Yaskawa INFORM job: cattua0.JBI

/JOB
//NAME cattua0
//POS
///NPOS 130,0,0,0,0,0
///TOOL 9
///POSTYPE PULSE
///PULSE
C00000=-149478,-3800,-72601,-72634,-83747,-23013
C00001=-158362,27238,-42051,-68147,-87155,-20871
C00002=-155378,40422,-20095,-70093,-86314,-22222
C00003=-152934,54036,4519,-71957,-85739,-23985
C00004=-152872,54426,5251,-72009,-85726,-24041
C00005=-152818,54830,6002,-72058,-85717,-24097
C00006=-152775,55247,6768,-72103,-85712,-24152
C00007=-152741,55675,7548,-72144,-85712,-24206
C00008=-152718,56112,8337,-72182,-85717,-24260
C00009=-152706,56556,9133,-72216,-85727,-24313
C00010=-152703,57006,9933,-72246,-85742,-24364
C00011=-152712,57461,10733,-72271,-85762,-24415
C00012=-152730,57917,11532,-72293,-85786,-24464
C00013=-152759,58374,12326,-72310,-85815,-24511
C00014=-152798,58830,13113,-72324,-85848,-24557
C00015=-152846,59283,13889,-72334,-85886,-24600
C00016=-152903,59731,14652,-72340,-85927,-24642
C00017=-152969,60172,15400,-72342,-85973,-24683
C00018=-153124,61027,16837,-72336,-86074,-24757
C00019=-153307,61842,18195,-72317,-86186,-24823
C00020=-153524,62645,19517,-72286,-86315,-24883
C00021=-153773,63424,20787,-72241,-86458,-24938
C00022=-154052,64166,21985,-72184,-86615,-24985
C00023=-154358,64860,23092,-72114,-86783,-25024
C00024=-154687,65495,24091,-72033,-86960,-25055
C00025=-155034,66063,24971,-71941,-87145,-25077
C00026=-155395,66557,25719,-71839,-87334,-25089
C00027=-156090,67486,27164,-71650,-87700,-25120
C00028=-156792,68395,28628,-71464,-88074,-25159
C00029=-157502,69283,30109,-71285,-88455,-25207
C00030=-158217,70146,31604,-71111,-88843,-25263
C00031=-158938,70984,33108,-70945,-89238,-25327
C00032=-159661,71794,34620,-70786,-89640,-25400
C00033=-160387,72575,36134,-70636,-90046,-25480
C00034=-161114,73326,37650,-70495,-90458,-25569
C00035=-161841,74047,39164,-70364,-90874,-25665
C00036=-162568,74735,40675,-70242,-91293,-25769
C00037=-163292,75392,42179,-70132,-91716,-25881
C00038=-164013,76015,43673,-70033,-92142,-25999
C00039=-164729,76606,45157,-69946,-92569,-26124
C00040=-165440,77164,46627,-69871,-92997,-26256
C00041=-166143,77688,48082,-69808,-93425,-26393
C00042=-166839,78181,49519,-69758,-93852,-26537
C00043=-167197,78385,50174,-69730,-94071,-26606
C00044=-167566,78510,50675,-69688,-94290,-26661
C00045=-167940,78553,51011,-69632,-94507,-26702
C00046=-168316,78512,51178,-69562,-94720,-26728
C00047=-168690,78390,51174,-69478,-94926,-26737
C00048=-169057,78191,51002,-69380,-95123,-26731
C00049=-169413,77920,50673,-69271,-95307,-26709
C00050=-169759,77583,50193,-69149,-95480,-26672
C00051=-170104,77167,49544,-69010,-95646,-26618
C00052=-170444,76676,48726,-68854,-95801,-26547
C00053=-170773,76114,47744,-68684,-95944,-26458
C00054=-170932,75809,47195,-68593,-96010,-26408
C00055=-171087,75489,46610,-68500,-96071,-26354
C00056=-171237,75156,45990,-68403,-96128,-26295
C00057=-171381,74810,45337,-68304,-96181,-26234
C00058=-171519,74454,44656,-68203,-96228,-26168
C00059=-171651,74088,43948,-68101,-96271,-26100
C00060=-171776,73715,43217,-67997,-96308,-26029
C00061=-171893,73336,42467,-67892,-96340,-25956
C00062=-172106,72568,40924,-67682,-96388,-25804
C00063=-176209,59482,15170,-63884,-97305,-23273
C00064=-180964,47935,-6371,-60041,-98451,-21150
C00065=-181093,47637,-6920,-59937,-98479,-21095
C00066=-181207,47321,-7519,-59832,-98497,-21036
C00067=-181305,46992,-8163,-59728,-98503,-20972
C00068=-181384,46655,-8839,-59627,-98496,-20905
C00069=-181443,46314,-9539,-59531,-98477,-20837
C00070=-181482,45976,-10249,-59441,-98446,-20767
C00071=-181498,45645,-10960,-59360,-98405,-20698
C00072=-181495,45326,-11657,-59288,-98354,-20632
C00073=-181473,45023,-12333,-59226,-98295,-20567
C00074=-181431,44725,-13010,-59171,-98226,-20504
C00075=-181369,44435,-13683,-59126,-98148,-20441
C00076=-181287,44157,-14341,-59090,-98061,-20381
C00077=-181186,43895,-14975,-59065,-97966,-20324
C00078=-181067,43652,-15576,-59051,-97865,-20271
C00079=-180931,43432,-16137,-59049,-97758,-20223
C00080=-180781,43237,-16651,-59058,-97649,-20180
C00081=-180331,42715,-18030,-59105,-97335,-20069
C00082=-179870,42191,-19389,-59167,-97022,-19965
C00083=-179397,41663,-20725,-59243,-96709,-19868
C00084=-178913,41133,-22039,-59333,-96396,-19778
C00085=-178417,40599,-23328,-59437,-96085,-19694
C00086=-177910,40063,-24592,-59555,-95774,-19618
C00087=-177391,39523,-25830,-59686,-95465,-19550
C00088=-176861,38981,-27041,-59831,-95157,-19488
C00089=-176321,38437,-28225,-59989,-94850,-19434
C00090=-175769,37891,-29380,-60160,-94545,-19387
C00091=-175207,37342,-30505,-60344,-94242,-19347
C00092=-174635,36792,-31599,-60540,-93941,-19315
C00093=-174053,36240,-32663,-60748,-93641,-19290
C00094=-173462,35687,-33694,-60968,-93344,-19272
C00095=-172862,35132,-34693,-61198,-93049,-19262
C00096=-172252,34577,-35659,-61440,-92755,-19259
C00097=-171634,34021,-36591,-61692,-92464,-19263
C00098=-171008,33464,-37488,-61954,-92175,-19274
C00099=-170375,32907,-38351,-62225,-91888,-19293
C00100=-169734,32350,-39178,-62506,-91604,-19319
C00101=-169086,31793,-39970,-62795,-91321,-19352
C00102=-168432,31237,-40725,-63091,-91041,-19392
C00103=-167773,30682,-41443,-63396,-90762,-19440
C00104=-167108,30129,-42124,-63707,-90486,-19494
C00105=-166440,29577,-42767,-64025,-90212,-19555
C00106=-165767,29028,-43372,-64348,-89940,-19622
C00107=-165092,28481,-43940,-64676,-89670,-19697
C00108=-164414,27937,-44469,-65009,-89403,-19777
C00109=-163734,27396,-44960,-65345,-89137,-19864
C00110=-163053,26860,-45412,-65685,-88873,-19957
C00111=-162372,26328,-45826,-66027,-88612,-20057
C00112=-161691,25800,-46202,-66371,-88352,-20162
C00113=-161451,25633,-46301,-66493,-88262,-20201
C00114=-161203,25495,-46349,-66621,-88168,-20243
C00115=-160950,25391,-46344,-66751,-88074,-20288
C00116=-160696,25322,-46286,-66884,-87981,-20335
C00117=-160444,25288,-46176,-67015,-87888,-20383
C00118=-160199,25292,-46016,-67145,-87798,-20431
C00119=-159962,25330,-45810,-67270,-87712,-20480
C00120=-159736,25403,-45562,-67390,-87631,-20527
C00121=-159515,25511,-45264,-67508,-87552,-20576
C00122=-159301,25658,-44916,-67623,-87476,-20624
C00123=-159099,25843,-44521,-67733,-87404,-20671
C00124=-158911,26064,-44083,-67836,-87338,-20717
C00125=-158741,26319,-43609,-67930,-87280,-20761
C00126=-158592,26603,-43106,-68014,-87229,-20801
C00127=-158465,26912,-42583,-68086,-87187,-20838
C00128=-158362,27238,-42051,-68147,-87155,-20871
C00129=-158362,19647,-34950,-70491,-88624,-24433
//INST
///DATE 2026/08/21 15:23
///COMM Generated using RoboDK
///ATTR SC,RW
///GROUP1 RB1
NOP
'Program generated by RoboDK v
'4.0.0 for Motoman UP50N on 21
'/08/2026 15:22:59
'Using nominal kinematics.
'Using Frame 2 (targets wrt ba
'se):
'-320.0,-1370.0,-236.0,0.0,0.0
',90.0
'Tool Teknomotor QTC C4147-C-D
'B Spindle should be close to:
'200.0,0.0,200.0,0.0,90.0,0.0
'Show Teknomotor QTC C4147-C-D
'B Spindle
DOUT OT#(9) ON
MOVJ C00000 VJ=10.00 PL=1
MOVL C00001 V=200.0 PL=1
MOVL C00002 V=60.0 PL=1
MOVL C00003 V=60.0 PL=1
MOVL C00004 V=60.0 PL=1
MOVL C00005 V=60.0 PL=1
MOVL C00006 V=60.0 PL=1
MOVL C00007 V=60.0 PL=1
MOVL C00008 V=60.0 PL=1
MOVL C00009 V=60.0 PL=1
MOVL C00010 V=60.0 PL=1
MOVL C00011 V=60.0 PL=1
MOVL C00012 V=60.0 PL=1
MOVL C00013 V=60.0 PL=1
MOVL C00014 V=60.0 PL=1
MOVL C00015 V=60.0 PL=1
MOVL C00016 V=60.0 PL=1
MOVL C00017 V=60.0 PL=1
MOVL C00018 V=60.0 PL=1
MOVL C00019 V=60.0 PL=1
MOVL C00020 V=60.0 PL=1
MOVL C00021 V=60.0 PL=1
MOVL C00022 V=60.0 PL=1
MOVL C00023 V=60.0 PL=1
MOVL C00024 V=60.0 PL=1
MOVL C00025 V=60.0 PL=1
MOVL C00026 V=60.0 PL=1
MOVL C00027 V=60.0 PL=1
MOVL C00028 V=60.0 PL=1
MOVL C00029 V=60.0 PL=1
MOVL C00030 V=60.0 PL=1
MOVL C00031 V=60.0 PL=1
MOVL C00032 V=60.0 PL=1
MOVL C00033 V=60.0 PL=1
MOVL C00034 V=60.0 PL=1
MOVL C00035 V=60.0 PL=1
MOVL C00036 V=60.0 PL=1
MOVL C00037 V=60.0 PL=1
MOVL C00038 V=60.0 PL=1
MOVL C00039 V=60.0 PL=1
MOVL C00040 V=60.0 PL=1
MOVL C00041 V=60.0 PL=1
MOVL C00042 V=60.0 PL=1
MOVL C00043 V=60.0 PL=1
MOVL C00044 V=60.0 PL=1
MOVL C00045 V=60.0 PL=1
MOVL C00046 V=60.0 PL=1
MOVL C00047 V=60.0 PL=1
MOVL C00048 V=60.0 PL=1
MOVL C00049 V=60.0 PL=1
MOVL C00050 V=60.0 PL=1
MOVL C00051 V=60.0 PL=1
MOVL C00052 V=60.0 PL=1
MOVL C00053 V=60.0 PL=1
MOVL C00054 V=60.0 PL=1
MOVL C00055 V=60.0 PL=1
MOVL C00056 V=60.0 PL=1
MOVL C00057 V=60.0 PL=1
MOVL C00058 V=60.0 PL=1
MOVL C00059 V=60.0 PL=1
MOVL C00060 V=60.0 PL=1
MOVL C00061 V=60.0 PL=1
MOVL C00062 V=60.0 PL=1
MOVL C00063 V=60.0 PL=1
MOVL C00064 V=60.0 PL=1
MOVL C00065 V=60.0 PL=1
MOVL C00066 V=60.0 PL=1
MOVL C00067 V=60.0 PL=1
MOVL C00068 V=60.0 PL=1
MOVL C00069 V=60.0 PL=1
MOVL C00070 V=60.0 PL=1
MOVL C00071 V=60.0 PL=1
MOVL C00072 V=60.0 PL=1
MOVL C00073 V=60.0 PL=1
MOVL C00074 V=60.0 PL=1
MOVL C00075 V=60.0 PL=1
MOVL C00076 V=60.0 PL=1
MOVL C00077 V=60.0 PL=1
MOVL C00078 V=60.0 PL=1
MOVL C00079 V=60.0 PL=1
MOVL C00080 V=60.0 PL=1
MOVL C00081 V=60.0 PL=1
MOVL C00082 V=60.0 PL=1
MOVL C00083 V=60.0 PL=1
MOVL C00084 V=60.0 PL=1
MOVL C00085 V=60.0 PL=1
MOVL C00086 V=60.0 PL=1
MOVL C00087 V=60.0 PL=1
MOVL C00088 V=60.0 PL=1
MOVL C00089 V=60.0 PL=1
MOVL C00090 V=60.0 PL=1
MOVL C00091 V=60.0 PL=1
MOVL C00092 V=60.0 PL=1
MOVL C00093 V=60.0 PL=1
MOVL C00094 V=60.0 PL=1
MOVL C00095 V=60.0 PL=1
MOVL C00096 V=60.0 PL=1
MOVL C00097 V=60.0 PL=1
MOVL C00098 V=60.0 PL=1
MOVL C00099 V=60.0 PL=1
MOVL C00100 V=60.0 PL=1
MOVL C00101 V=60.0 PL=1
MOVL C00102 V=60.0 PL=1
MOVL C00103 V=60.0 PL=1
MOVL C00104 V=60.0 PL=1
MOVL C00105 V=60.0 PL=1
MOVL C00106 V=60.0 PL=1
MOVL C00107 V=60.0 PL=1
MOVL C00108 V=60.0 PL=1
MOVL C00109 V=60.0 PL=1
MOVL C00110 V=60.0 PL=1
MOVL C00111 V=60.0 PL=1
MOVL C00112 V=60.0 PL=1
MOVL C00113 V=60.0 PL=1
MOVL C00114 V=60.0 PL=1
MOVL C00115 V=60.0 PL=1
MOVL C00116 V=60.0 PL=1
MOVL C00117 V=60.0 PL=1
MOVL C00118 V=60.0 PL=1
MOVL C00119 V=60.0 PL=1
MOVL C00120 V=60.0 PL=1
MOVL C00121 V=60.0 PL=1
MOVL C00122 V=60.0 PL=1
MOVL C00123 V=60.0 PL=1
MOVL C00124 V=60.0 PL=1
MOVL C00125 V=60.0 PL=1
MOVL C00126 V=60.0 PL=1
MOVL C00127 V=60.0 PL=1
MOVL C00128 V=60.0 PL=1
MOVL C00129 V=200.0 PL=1
DOUT OT#(9) OFF
END
